(* IEC 61131-3 sources: VLSI-SoC2026-SoftPLC-Paper/openplc/test_C_modularity/pous/functions, 1 file *)

(* ---- ClampInt.st ---- *)
FUNCTION ClampInt : INT
VAR_INPUT
    x : INT;
    minVal : INT;
    maxVal : INT;
END_VAR

IF x < minVal THEN
    ClampInt := minVal;
ELSIF x > maxVal THEN
    ClampInt := maxVal;
ELSE
    ClampInt := x;
END_IF;

END_FUNCTION
